% RSLogix 500 project MILLIH2O.RSS, saved by version 12.00.00.00 %
PROJECT "MILLIH2O"    % processor: MicroLogix 1400 %

PROGRAM FILES
  LAD 2   13 rungs
  LAD 3   41 rungs
  LAD 4   59 rungs
  LAD 5   7 rungs
  LAD 6   5 rungs
  LAD 7   8 rungs
  LAD 8   86 rungs

DATA FILES
  O0 OUTPUT  8 elements
  I1 INPUT  8 elements
  S2 STATUS  66 elements
  B3 BINARY  20 elements
  T4 TIMER  27 elements
  C5 COUNTER  11 elements
  R6 CONTROL  1 elements
  N7 INTEGER  50 elements
  F8 FLOAT  133 elements
  N9   17 elements
  F10   3 elements
  B11   5 elements
  F12   23 elements
  N13   50 elements
  N14   4 elements
  C15   10 elements
  C16   10 elements
  B17   4 elements
  F18   60 elements
  F19   10 elements
  N20   100 elements
  B25   1 elements
  B26   1 elements
  F28   10 elements

LADDER 2
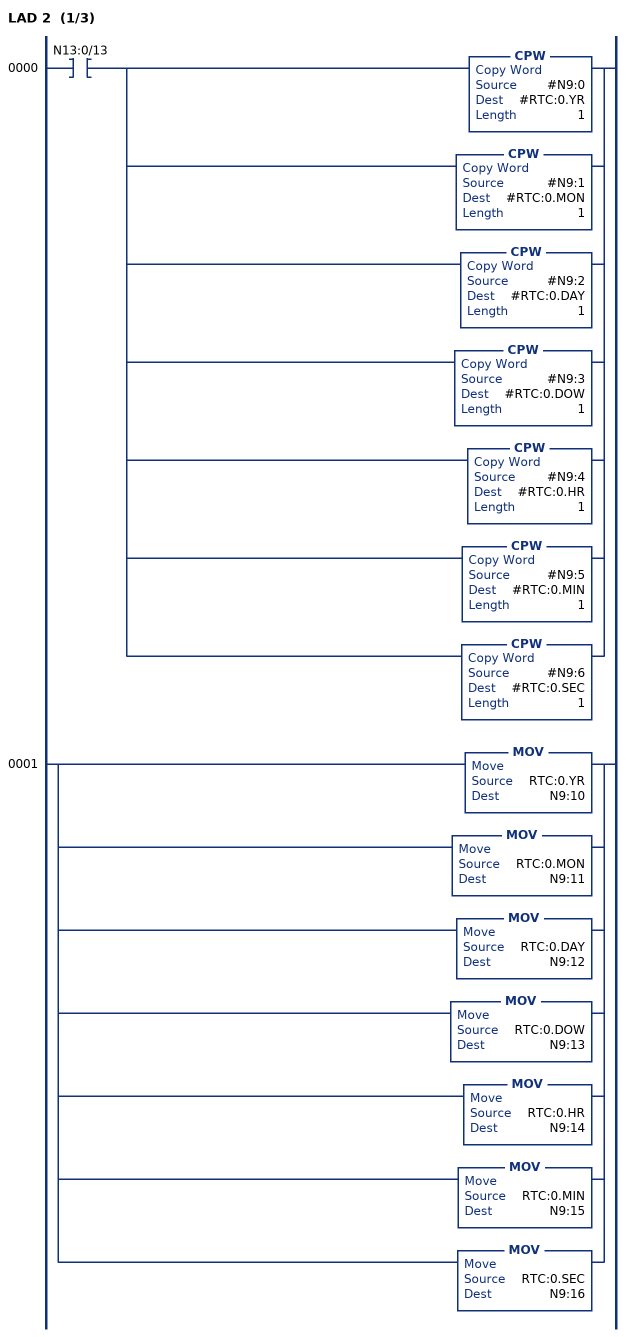
% Rung: 0 %
SOR XIC N13:0/13 BST CPW #N9:0 #RTC:0.YR 1 NXB CPW #N9:1 #RTC:0.MON 1 NXB CPW #N9:2 #RTC:0.DAY 1 NXB CPW #N9:3 #RTC:0.DOW 1 NXB CPW #N9:4 #RTC:0.HR 1 NXB CPW #N9:5 #RTC:0.MIN 1 NXB CPW #N9:6 #RTC:0.SEC 1 BND EOR
% Rung: 1 %
SOR BST MOV RTC:0.YR N9:10 NXB MOV RTC:0.MON N9:11 NXB MOV RTC:0.DAY N9:12 NXB MOV RTC:0.DOW N9:13 NXB MOV RTC:0.HR N9:14 NXB MOV RTC:0.MIN N9:15 NXB MOV RTC:0.SEC N9:16 BND EOR

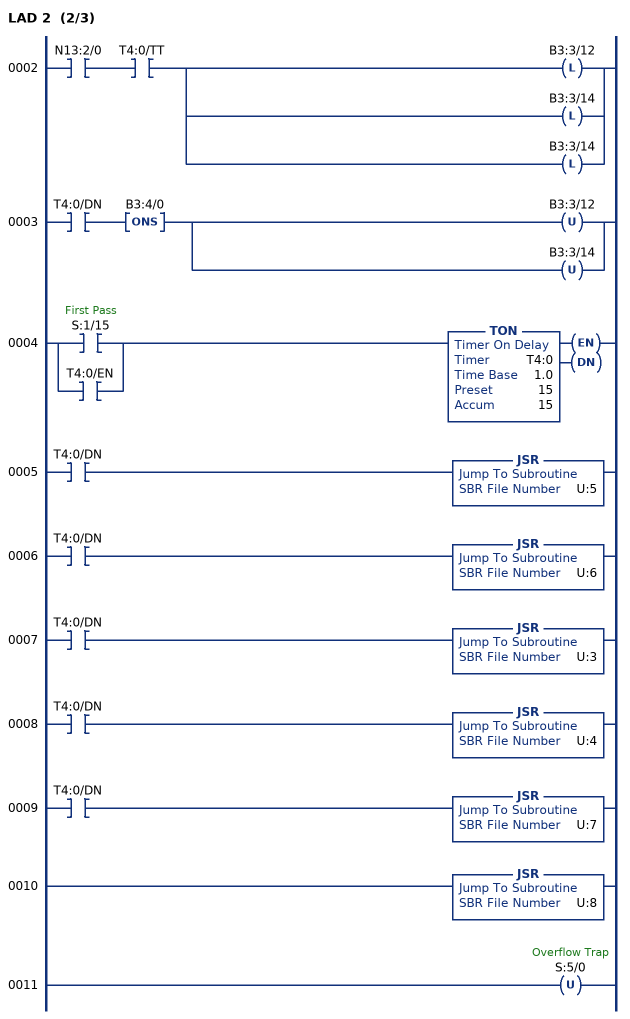
% Rung: 2 %
SOR XIC N13:2/0 XIC T4:0/TT BST OTL B3:3/12 NXB OTL B3:3/14 NXB OTL B3:3/14 BND EOR
% Rung: 3 %
SOR XIC T4:0/DN ONS B3:4/0 BST OTU B3:3/12 NXB OTU B3:3/14 BND EOR
% Rung: 4 %
SOR BST XIC S:1/15 NXB XIC T4:0/EN BND TON T4:0 1.0 15 15 EOR
%   S:1/15  "First Pass" %
% Rung: 5 %
SOR XIC T4:0/DN JSR U:5 EOR
% Rung: 6 %
SOR XIC T4:0/DN JSR U:6 EOR
% Rung: 7 %
SOR XIC T4:0/DN JSR U:3 EOR
% Rung: 8 %
SOR XIC T4:0/DN JSR U:4 EOR
% Rung: 9 %
SOR XIC T4:0/DN JSR U:7 EOR
% Rung: 10 %
SOR JSR U:8 EOR
% Rung: 11 %
SOR OTU S:5/0 EOR
%   S:5/0  "Overflow Trap" %

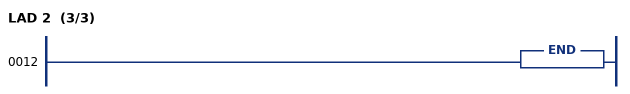
% Rung: 12 %
SOR END EOR

LADDER 3
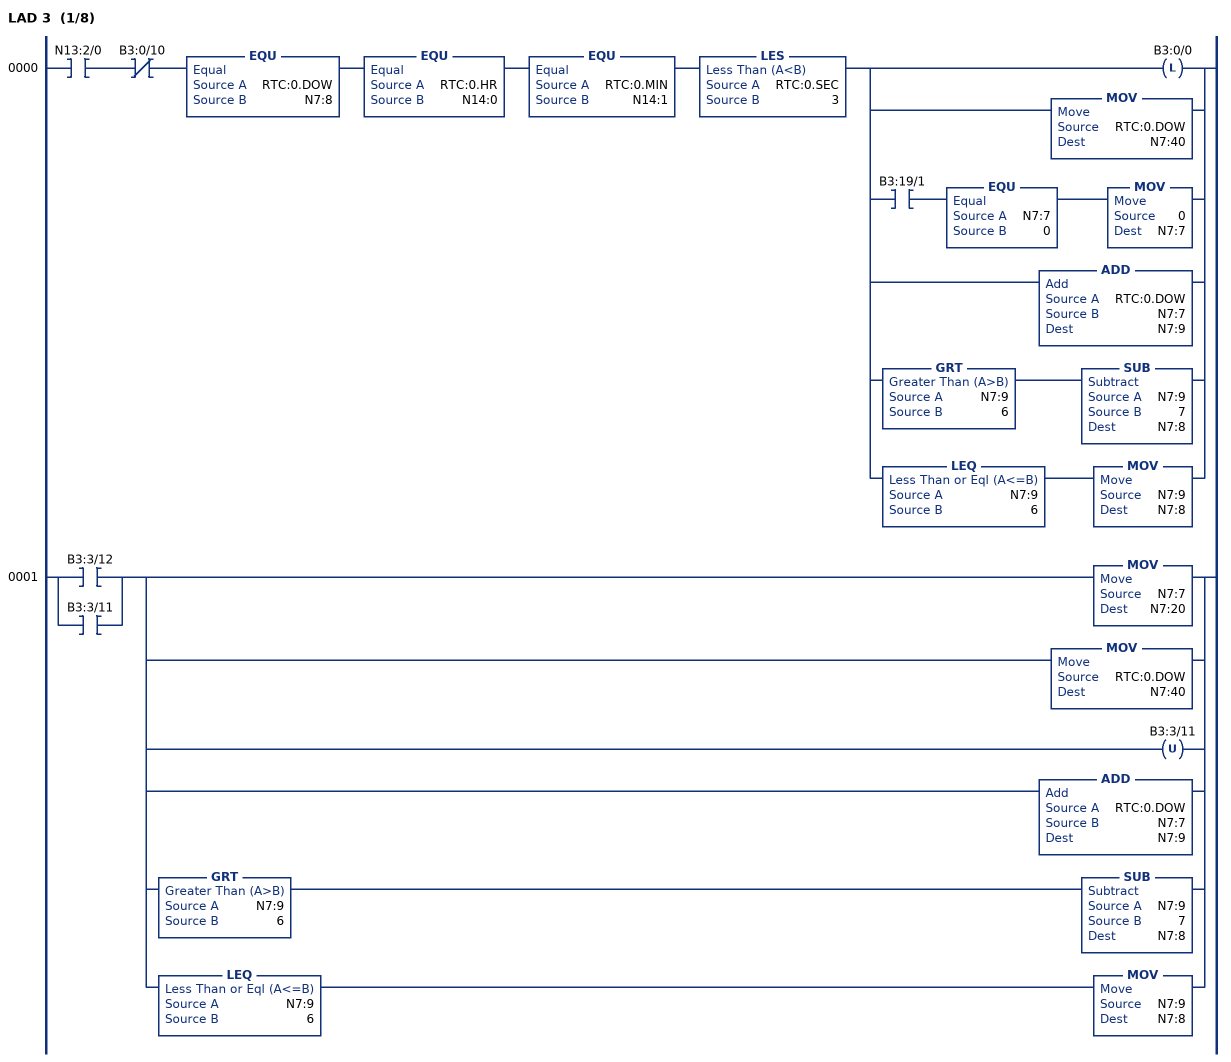
% Rung: 0 %
SOR XIC N13:2/0 XIO B3:0/10 EQU RTC:0.DOW N7:8 EQU RTC:0.HR N14:0 EQU RTC:0.MIN N14:1 LES RTC:0.SEC 3 BST OTL B3:0/0 NXB MOV RTC:0.DOW N7:40 NXB XIC B3:19/1 EQU N7:7 0 MOV 0 N7:7 NXB ADD RTC:0.DOW N7:7 N7:9 NXB GRT N7:9 6 SUB N7:9 7 N7:8 NXB LEQ N7:9 6 MOV N7:9 N7:8 BND EOR
% Rung: 1 %
SOR BST XIC B3:3/12 NXB XIC B3:3/11 BND BST MOV N7:7 N7:20 NXB MOV RTC:0.DOW N7:40 NXB OTU B3:3/11 NXB ADD RTC:0.DOW N7:7 N7:9 NXB GRT N7:9 6 SUB N7:9 7 N7:8 NXB LEQ N7:9 6 MOV N7:9 N7:8 BND EOR

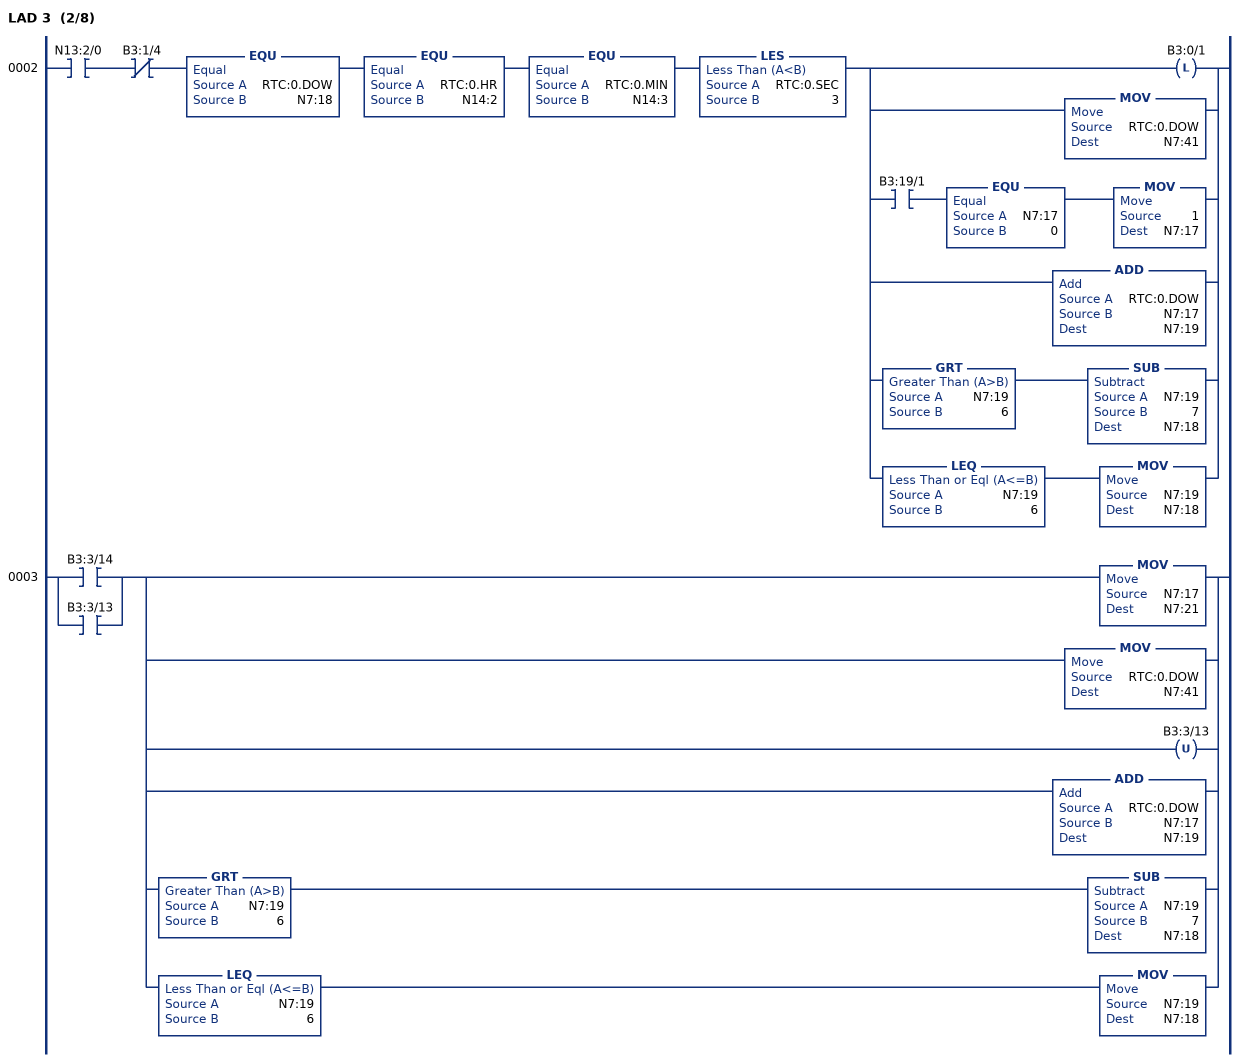
% Rung: 2 %
SOR XIC N13:2/0 XIO B3:1/4 EQU RTC:0.DOW N7:18 EQU RTC:0.HR N14:2 EQU RTC:0.MIN N14:3 LES RTC:0.SEC 3 BST OTL B3:0/1 NXB MOV RTC:0.DOW N7:41 NXB XIC B3:19/1 EQU N7:17 0 MOV 1 N7:17 NXB ADD RTC:0.DOW N7:17 N7:19 NXB GRT N7:19 6 SUB N7:19 7 N7:18 NXB LEQ N7:19 6 MOV N7:19 N7:18 BND EOR
% Rung: 3 %
SOR BST XIC B3:3/14 NXB XIC B3:3/13 BND BST MOV N7:17 N7:21 NXB MOV RTC:0.DOW N7:41 NXB OTU B3:3/13 NXB ADD RTC:0.DOW N7:17 N7:19 NXB GRT N7:19 6 SUB N7:19 7 N7:18 NXB LEQ N7:19 6 MOV N7:19 N7:18 BND EOR

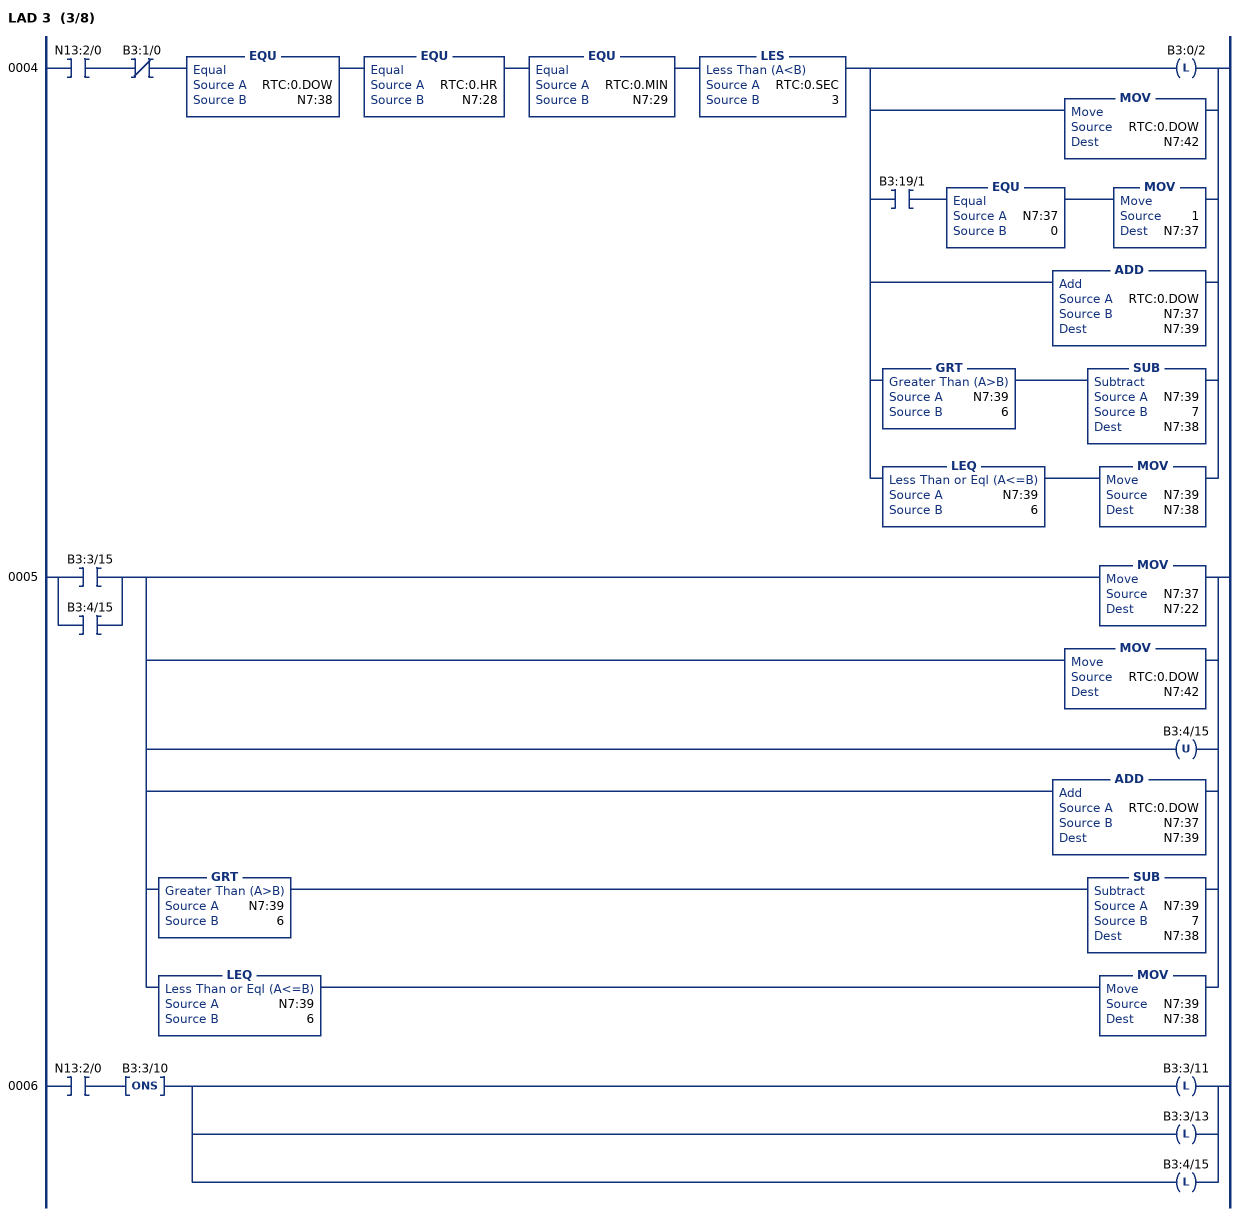
% Rung: 4 %
SOR XIC N13:2/0 XIO B3:1/0 EQU RTC:0.DOW N7:38 EQU RTC:0.HR N7:28 EQU RTC:0.MIN N7:29 LES RTC:0.SEC 3 BST OTL B3:0/2 NXB MOV RTC:0.DOW N7:42 NXB XIC B3:19/1 EQU N7:37 0 MOV 1 N7:37 NXB ADD RTC:0.DOW N7:37 N7:39 NXB GRT N7:39 6 SUB N7:39 7 N7:38 NXB LEQ N7:39 6 MOV N7:39 N7:38 BND EOR
% Rung: 5 %
SOR BST XIC B3:3/15 NXB XIC B3:4/15 BND BST MOV N7:37 N7:22 NXB MOV RTC:0.DOW N7:42 NXB OTU B3:4/15 NXB ADD RTC:0.DOW N7:37 N7:39 NXB GRT N7:39 6 SUB N7:39 7 N7:38 NXB LEQ N7:39 6 MOV N7:39 N7:38 BND EOR
% Rung: 6 %
SOR XIC N13:2/0 ONS B3:3/10 BST OTL B3:3/11 NXB OTL B3:3/13 NXB OTL B3:4/15 BND EOR

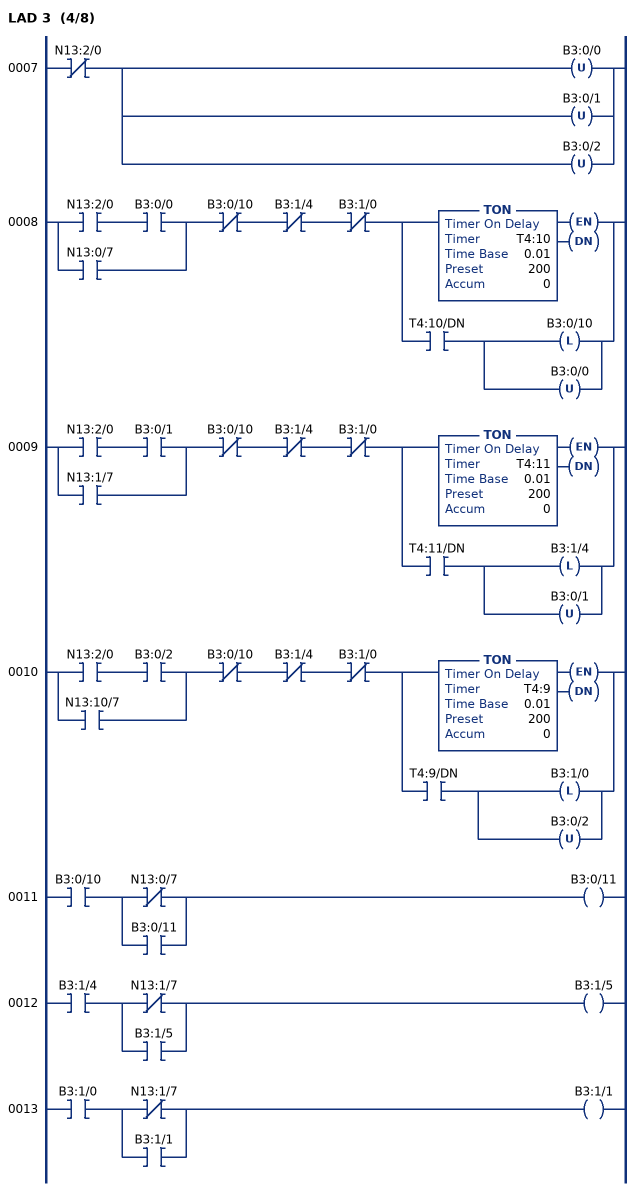
% Rung: 7 %
SOR XIO N13:2/0 BST OTU B3:0/0 NXB OTU B3:0/1 NXB OTU B3:0/2 BND EOR
% Rung: 8 %
SOR BST XIC N13:2/0 XIC B3:0/0 NXB XIC N13:0/7 BND XIO B3:0/10 XIO B3:1/4 XIO B3:1/0 BST TON T4:10 0.01 200 0 NXB XIC T4:10/DN BST OTL B3:0/10 NXB OTU B3:0/0 BND BND EOR
% Rung: 9 %
SOR BST XIC N13:2/0 XIC B3:0/1 NXB XIC N13:1/7 BND XIO B3:0/10 XIO B3:1/4 XIO B3:1/0 BST TON T4:11 0.01 200 0 NXB XIC T4:11/DN BST OTL B3:1/4 NXB OTU B3:0/1 BND BND EOR
% Rung: 10 %
SOR BST XIC N13:2/0 XIC B3:0/2 NXB XIC N13:10/7 BND XIO B3:0/10 XIO B3:1/4 XIO B3:1/0 BST TON T4:9 0.01 200 0 NXB XIC T4:9/DN BST OTL B3:1/0 NXB OTU B3:0/2 BND BND EOR
% Rung: 11 %
SOR XIC B3:0/10 BST XIO N13:0/7 NXB XIC B3:0/11 BND OTE B3:0/11 EOR
% Rung: 12 %
SOR XIC B3:1/4 BST XIO N13:1/7 NXB XIC B3:1/5 BND OTE B3:1/5 EOR
% Rung: 13 %
SOR XIC B3:1/0 BST XIO N13:1/7 NXB XIC B3:1/1 BND OTE B3:1/1 EOR

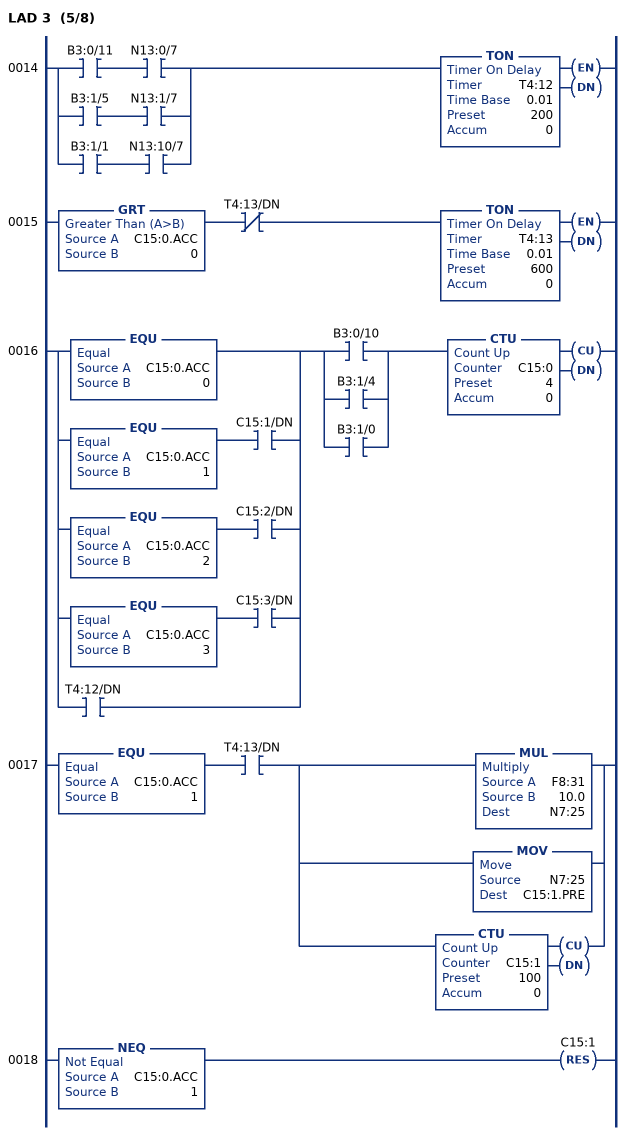
% Rung: 14 %
SOR BST XIC B3:0/11 XIC N13:0/7 NXB XIC B3:1/5 XIC N13:1/7 NXB XIC B3:1/1 XIC N13:10/7 BND TON T4:12 0.01 200 0 EOR
% Rung: 15 %
SOR GRT C15:0.ACC 0 XIO T4:13/DN TON T4:13 0.01 600 0 EOR
% Rung: 16 %
SOR BST EQU C15:0.ACC 0 NXB EQU C15:0.ACC 1 XIC C15:1/DN NXB EQU C15:0.ACC 2 XIC C15:2/DN NXB EQU C15:0.ACC 3 XIC C15:3/DN NXB XIC T4:12/DN BND BST XIC B3:0/10 NXB XIC B3:1/4 NXB XIC B3:1/0 BND CTU C15:0 4 0 EOR
% Rung: 17 %
SOR EQU C15:0.ACC 1 XIC T4:13/DN BST MUL F8:31 10.0 N7:25 NXB MOV N7:25 C15:1.PRE NXB CTU C15:1 100 0 BND EOR
% Rung: 18 %
SOR NEQ C15:0.ACC 1 RES C15:1 EOR

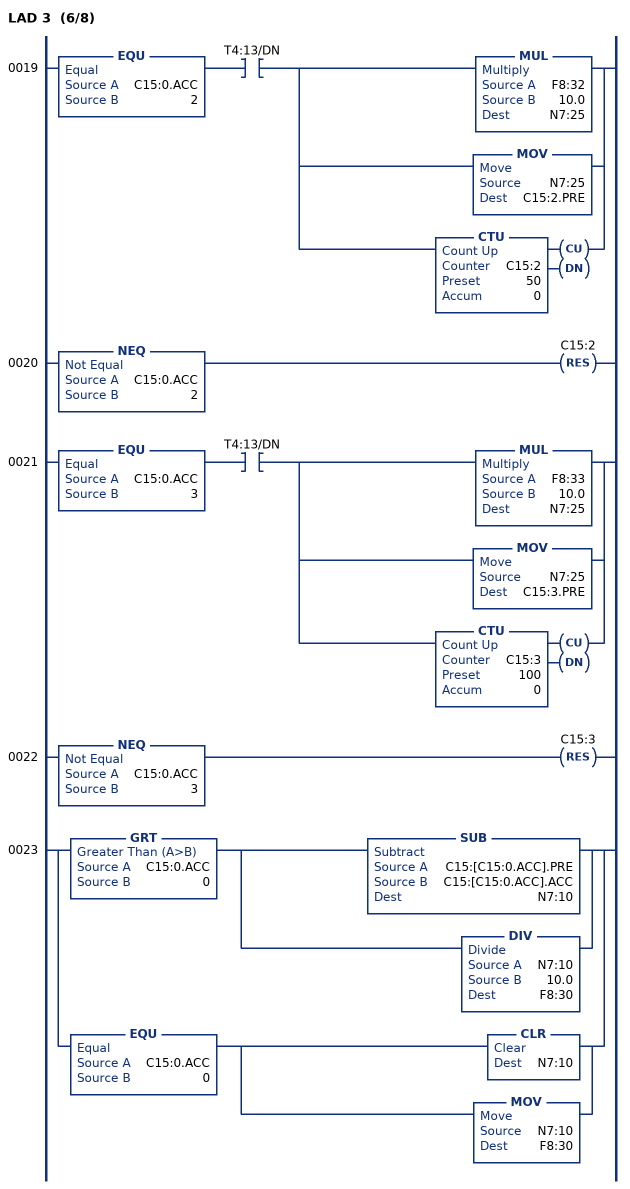
% Rung: 19 %
SOR EQU C15:0.ACC 2 XIC T4:13/DN BST MUL F8:32 10.0 N7:25 NXB MOV N7:25 C15:2.PRE NXB CTU C15:2 50 0 BND EOR
% Rung: 20 %
SOR NEQ C15:0.ACC 2 RES C15:2 EOR
% Rung: 21 %
SOR EQU C15:0.ACC 3 XIC T4:13/DN BST MUL F8:33 10.0 N7:25 NXB MOV N7:25 C15:3.PRE NXB CTU C15:3 100 0 BND EOR
% Rung: 22 %
SOR NEQ C15:0.ACC 3 RES C15:3 EOR
% Rung: 23 %
SOR BST GRT C15:0.ACC 0 BST SUB C15:[C15:0.ACC].PRE C15:[C15:0.ACC].ACC N7:10 NXB DIV N7:10 10.0 F8:30 BND NXB EQU C15:0.ACC 0 BST CLR N7:10 NXB MOV N7:10 F8:30 BND BND EOR

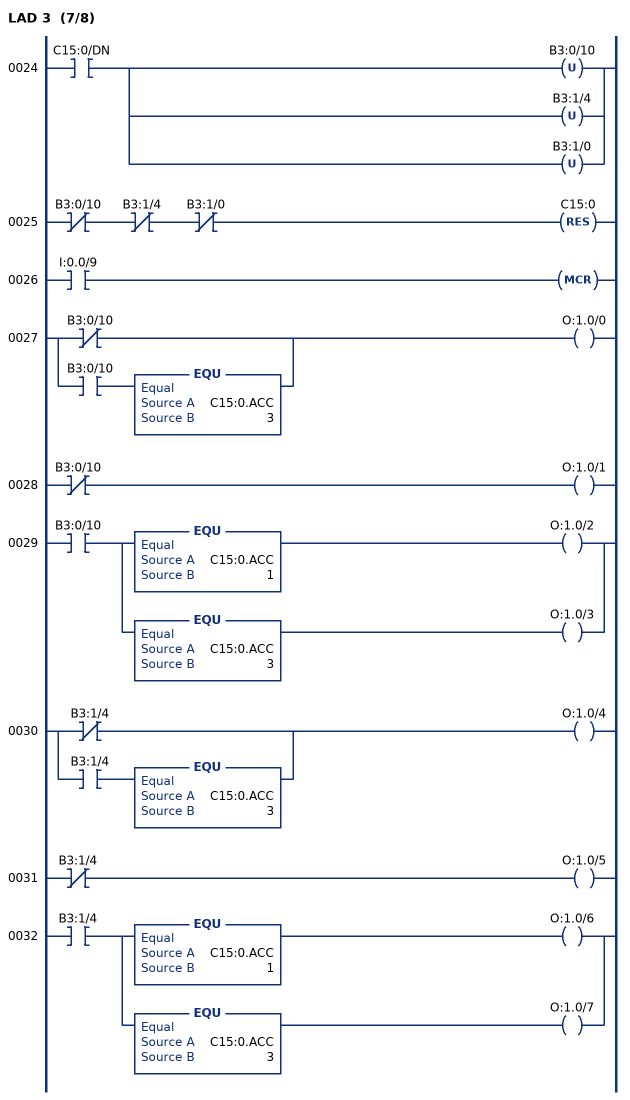
% Rung: 24 %
SOR XIC C15:0/DN BST OTU B3:0/10 NXB OTU B3:1/4 NXB OTU B3:1/0 BND EOR
% Rung: 25 %
SOR XIO B3:0/10 XIO B3:1/4 XIO B3:1/0 RES C15:0 EOR
% Rung: 26 %
SOR XIC I:0.0/9 MCR EOR
% Rung: 27 %
SOR BST XIO B3:0/10 NXB XIC B3:0/10 EQU C15:0.ACC 3 BND OTE O:1.0/0 EOR
% Rung: 28 %
SOR XIO B3:0/10 OTE O:1.0/1 EOR
% Rung: 29 %
SOR XIC B3:0/10 BST EQU C15:0.ACC 1 OTE O:1.0/2 NXB EQU C15:0.ACC 3 OTE O:1.0/3 BND EOR
% Rung: 30 %
SOR BST XIO B3:1/4 NXB XIC B3:1/4 EQU C15:0.ACC 3 BND OTE O:1.0/4 EOR
% Rung: 31 %
SOR XIO B3:1/4 OTE O:1.0/5 EOR
% Rung: 32 %
SOR XIC B3:1/4 BST EQU C15:0.ACC 1 OTE O:1.0/6 NXB EQU C15:0.ACC 3 OTE O:1.0/7 BND EOR

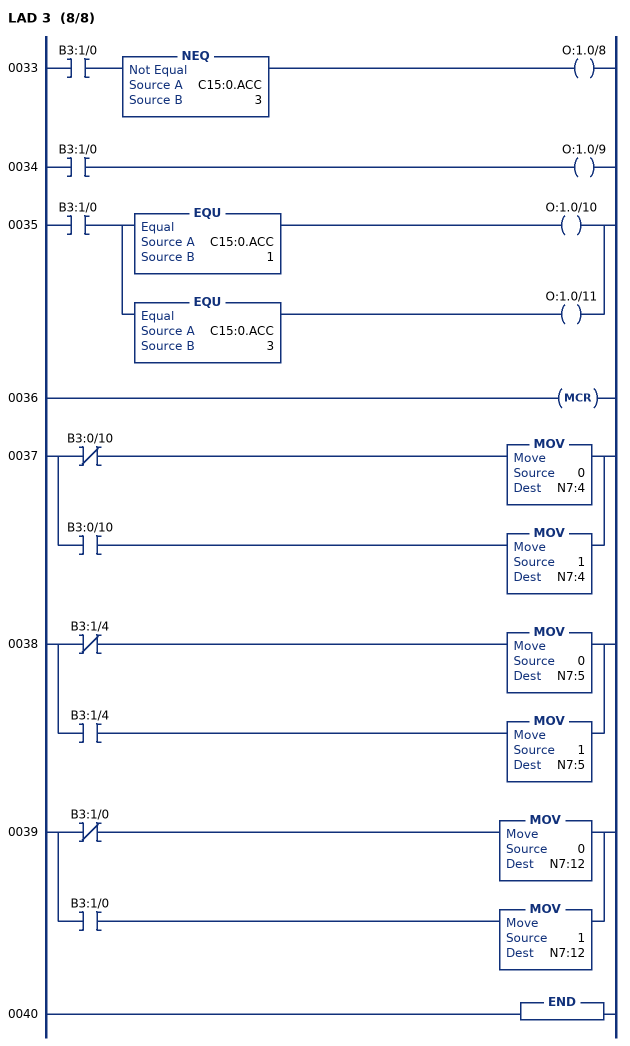
% Rung: 33 %
SOR XIC B3:1/0 NEQ C15:0.ACC 3 OTE O:1.0/8 EOR
% Rung: 34 %
SOR XIC B3:1/0 OTE O:1.0/9 EOR
% Rung: 35 %
SOR XIC B3:1/0 BST EQU C15:0.ACC 1 OTE O:1.0/10 NXB EQU C15:0.ACC 3 OTE O:1.0/11 BND EOR
% Rung: 36 %
SOR MCR EOR
% Rung: 37 %
SOR BST XIO B3:0/10 MOV 0 N7:4 NXB XIC B3:0/10 MOV 1 N7:4 BND EOR
% Rung: 38 %
SOR BST XIO B3:1/4 MOV 0 N7:5 NXB XIC B3:1/4 MOV 1 N7:5 BND EOR
% Rung: 39 %
SOR BST XIO B3:1/0 MOV 0 N7:12 NXB XIC B3:1/0 MOV 1 N7:12 BND EOR
% Rung: 40 %
SOR END EOR

LADDER 4
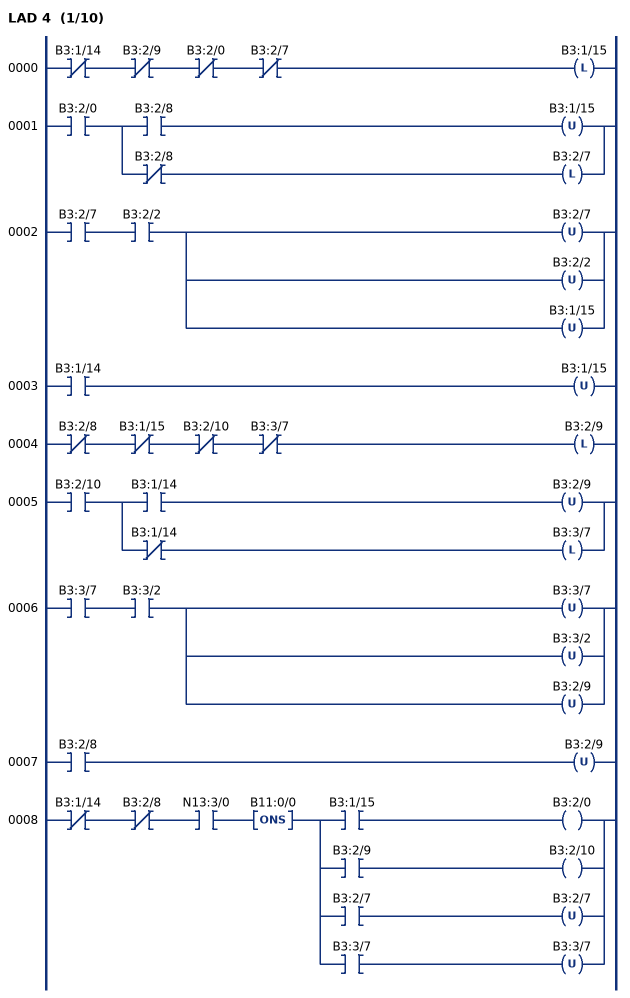
% Rung: 0 %
SOR XIO B3:1/14 XIO B3:2/9 XIO B3:2/0 XIO B3:2/7 OTL B3:1/15 EOR
% Rung: 1 %
SOR XIC B3:2/0 BST XIC B3:2/8 OTU B3:1/15 NXB XIO B3:2/8 OTL B3:2/7 BND EOR
% Rung: 2 %
SOR XIC B3:2/7 XIC B3:2/2 BST OTU B3:2/7 NXB OTU B3:2/2 NXB OTU B3:1/15 BND EOR
% Rung: 3 %
SOR XIC B3:1/14 OTU B3:1/15 EOR
% Rung: 4 %
SOR XIO B3:2/8 XIO B3:1/15 XIO B3:2/10 XIO B3:3/7 OTL B3:2/9 EOR
% Rung: 5 %
SOR XIC B3:2/10 BST XIC B3:1/14 OTU B3:2/9 NXB XIO B3:1/14 OTL B3:3/7 BND EOR
% Rung: 6 %
SOR XIC B3:3/7 XIC B3:3/2 BST OTU B3:3/7 NXB OTU B3:3/2 NXB OTU B3:2/9 BND EOR
% Rung: 7 %
SOR XIC B3:2/8 OTU B3:2/9 EOR
% Rung: 8 %
SOR XIO B3:1/14 XIO B3:2/8 XIC N13:3/0 ONS B11:0/0 BST XIC B3:1/15 OTE B3:2/0 NXB XIC B3:2/9 OTE B3:2/10 NXB XIC B3:2/7 OTU B3:2/7 NXB XIC B3:3/7 OTU B3:3/7 BND EOR

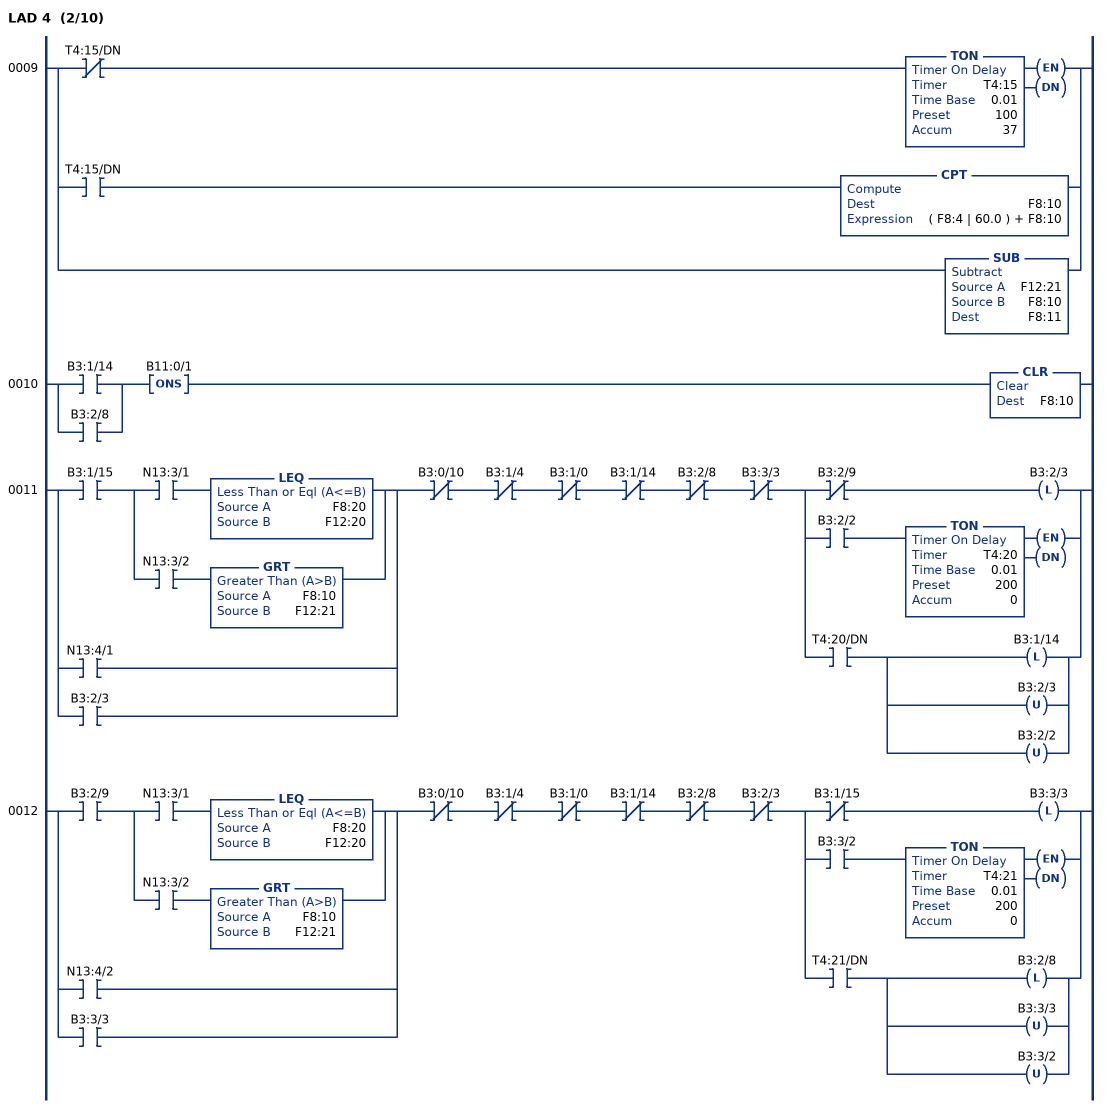
% Rung: 9 %
SOR BST XIO T4:15/DN TON T4:15 0.01 100 37 NXB XIC T4:15/DN CPT F8:10 " ( F8:4 | 60.0 ) + F8:10 " NXB SUB F12:21 F8:10 F8:11 BND EOR
% Rung: 10 %
SOR BST XIC B3:1/14 NXB XIC B3:2/8 BND ONS B11:0/1 CLR F8:10 EOR
% Rung: 11 %
SOR BST XIC B3:1/15 BST XIC N13:3/1 LEQ F8:20 F12:20 NXB XIC N13:3/2 GRT F8:10 F12:21 BND NXB XIC N13:4/1 NXB XIC B3:2/3 BND XIO B3:0/10 XIO B3:1/4 XIO B3:1/0 XIO B3:1/14 XIO B3:2/8 XIO B3:3/3 BST XIO B3:2/9 OTL B3:2/3 NXB XIC B3:2/2 TON T4:20 0.01 200 0 NXB XIC T4:20/DN BST OTL B3:1/14 NXB OTU B3:2/3 NXB OTU B3:2/2 BND BND EOR
% Rung: 12 %
SOR BST XIC B3:2/9 BST XIC N13:3/1 LEQ F8:20 F12:20 NXB XIC N13:3/2 GRT F8:10 F12:21 BND NXB XIC N13:4/2 NXB XIC B3:3/3 BND XIO B3:0/10 XIO B3:1/4 XIO B3:1/0 XIO B3:1/14 XIO B3:2/8 XIO B3:2/3 BST XIO B3:1/15 OTL B3:3/3 NXB XIC B3:3/2 TON T4:21 0.01 200 0 NXB XIC T4:21/DN BST OTL B3:2/8 NXB OTU B3:3/3 NXB OTU B3:3/2 BND BND EOR

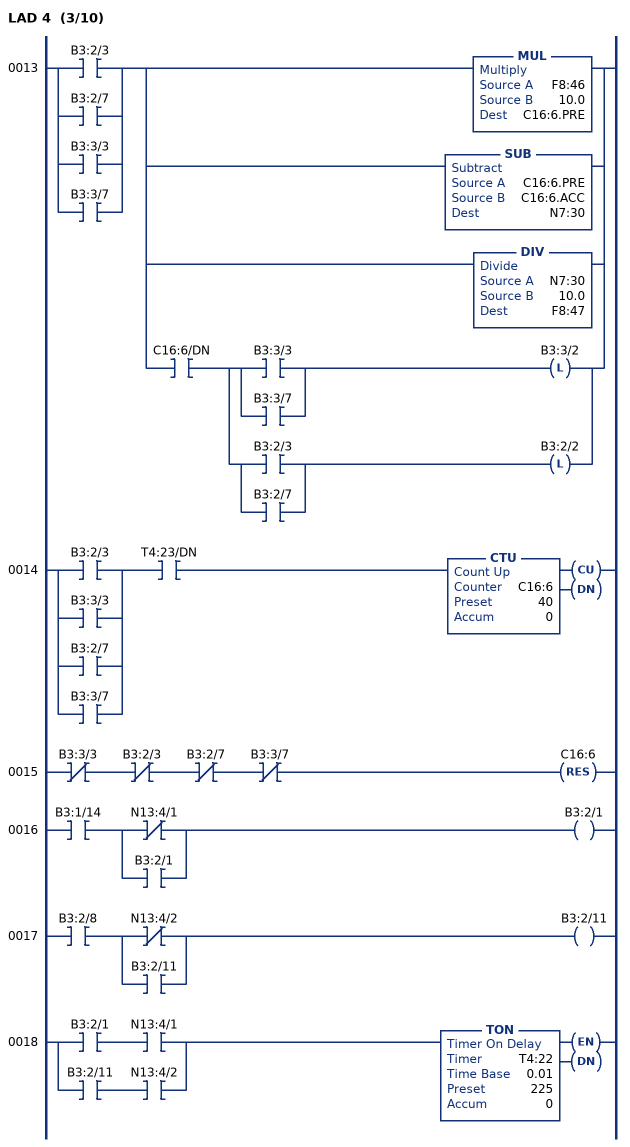
% Rung: 13 %
SOR BST XIC B3:2/3 NXB XIC B3:2/7 NXB XIC B3:3/3 NXB XIC B3:3/7 BND BST MUL F8:46 10.0 C16:6.PRE NXB SUB C16:6.PRE C16:6.ACC N7:30 NXB DIV N7:30 10.0 F8:47 NXB XIC C16:6/DN BST BST XIC B3:3/3 NXB XIC B3:3/7 BND OTL B3:3/2 NXB BST XIC B3:2/3 NXB XIC B3:2/7 BND OTL B3:2/2 BND BND EOR
% Rung: 14 %
SOR BST XIC B3:2/3 NXB XIC B3:3/3 NXB XIC B3:2/7 NXB XIC B3:3/7 BND XIC T4:23/DN CTU C16:6 40 0 EOR
% Rung: 15 %
SOR XIO B3:3/3 XIO B3:2/3 XIO B3:2/7 XIO B3:3/7 RES C16:6 EOR
% Rung: 16 %
SOR XIC B3:1/14 BST XIO N13:4/1 NXB XIC B3:2/1 BND OTE B3:2/1 EOR
% Rung: 17 %
SOR XIC B3:2/8 BST XIO N13:4/2 NXB XIC B3:2/11 BND OTE B3:2/11 EOR
% Rung: 18 %
SOR BST XIC B3:2/1 XIC N13:4/1 NXB XIC B3:2/11 XIC N13:4/2 BND TON T4:22 0.01 225 0 EOR

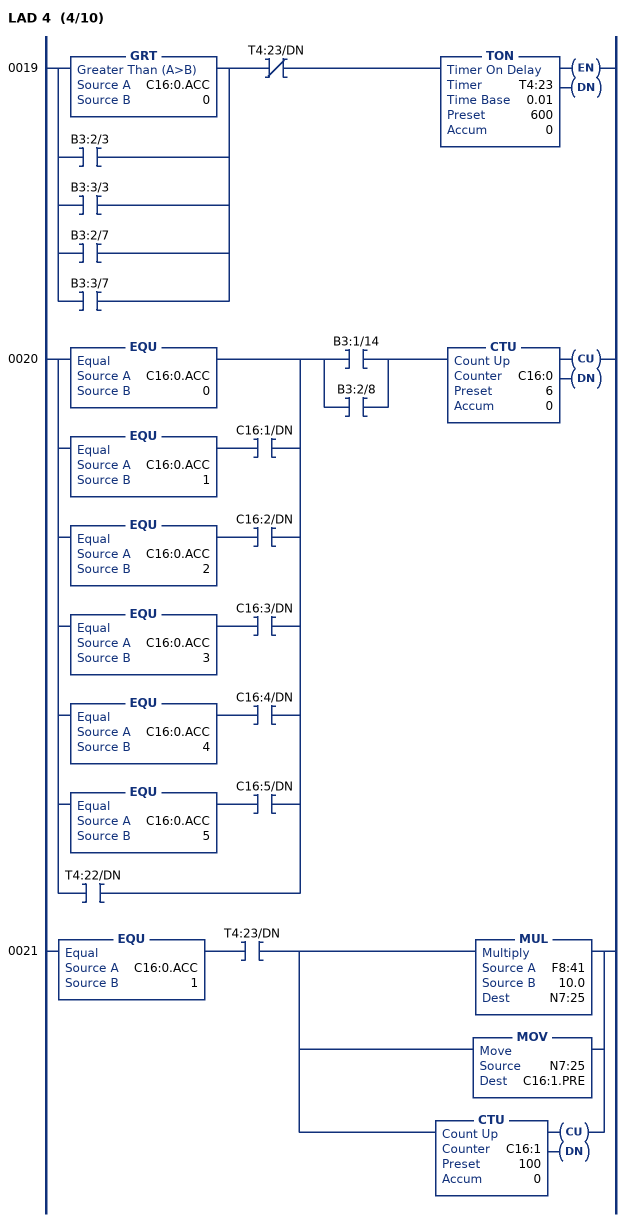
% Rung: 19 %
SOR BST GRT C16:0.ACC 0 NXB XIC B3:2/3 NXB XIC B3:3/3 NXB XIC B3:2/7 NXB XIC B3:3/7 BND XIO T4:23/DN TON T4:23 0.01 600 0 EOR
% Rung: 20 %
SOR BST EQU C16:0.ACC 0 NXB EQU C16:0.ACC 1 XIC C16:1/DN NXB EQU C16:0.ACC 2 XIC C16:2/DN NXB EQU C16:0.ACC 3 XIC C16:3/DN NXB EQU C16:0.ACC 4 XIC C16:4/DN NXB EQU C16:0.ACC 5 XIC C16:5/DN NXB XIC T4:22/DN BND BST XIC B3:1/14 NXB XIC B3:2/8 BND CTU C16:0 6 0 EOR
% Rung: 21 %
SOR EQU C16:0.ACC 1 XIC T4:23/DN BST MUL F8:41 10.0 N7:25 NXB MOV N7:25 C16:1.PRE NXB CTU C16:1 100 0 BND EOR

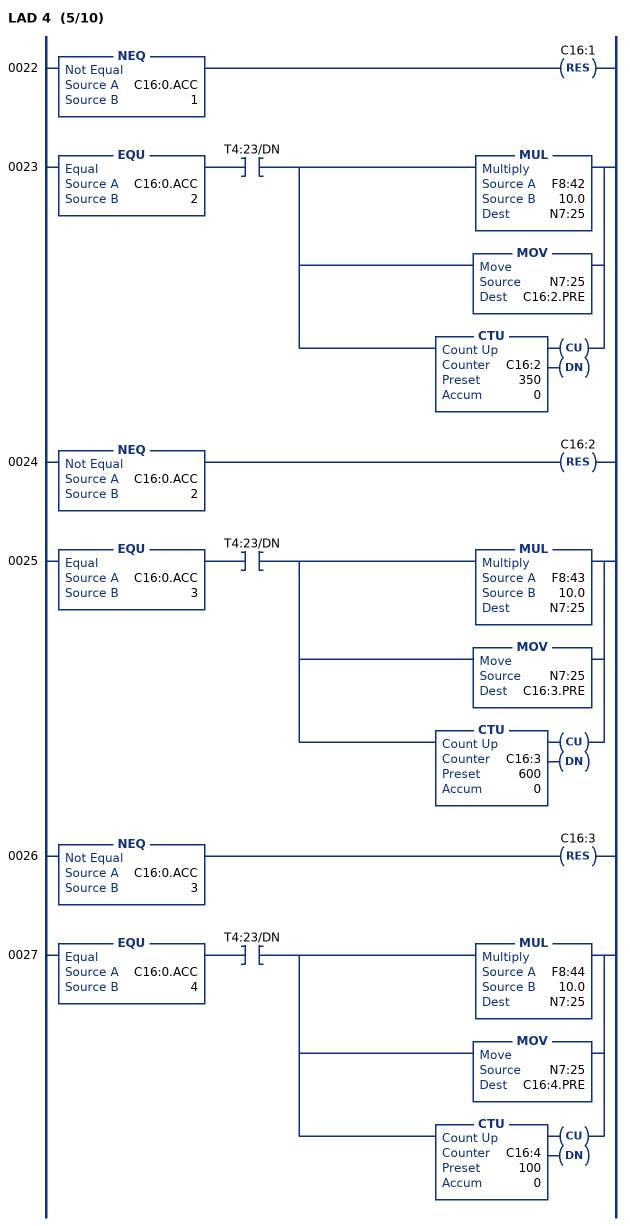
% Rung: 22 %
SOR NEQ C16:0.ACC 1 RES C16:1 EOR
% Rung: 23 %
SOR EQU C16:0.ACC 2 XIC T4:23/DN BST MUL F8:42 10.0 N7:25 NXB MOV N7:25 C16:2.PRE NXB CTU C16:2 350 0 BND EOR
% Rung: 24 %
SOR NEQ C16:0.ACC 2 RES C16:2 EOR
% Rung: 25 %
SOR EQU C16:0.ACC 3 XIC T4:23/DN BST MUL F8:43 10.0 N7:25 NXB MOV N7:25 C16:3.PRE NXB CTU C16:3 600 0 BND EOR
% Rung: 26 %
SOR NEQ C16:0.ACC 3 RES C16:3 EOR
% Rung: 27 %
SOR EQU C16:0.ACC 4 XIC T4:23/DN BST MUL F8:44 10.0 N7:25 NXB MOV N7:25 C16:4.PRE NXB CTU C16:4 100 0 BND EOR

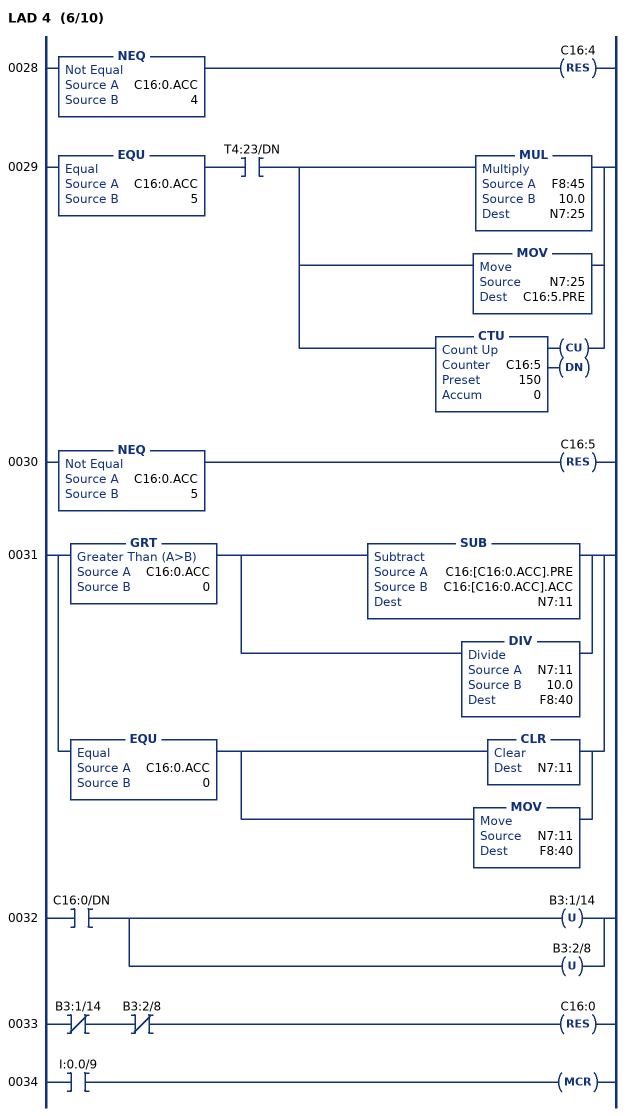
% Rung: 28 %
SOR NEQ C16:0.ACC 4 RES C16:4 EOR
% Rung: 29 %
SOR EQU C16:0.ACC 5 XIC T4:23/DN BST MUL F8:45 10.0 N7:25 NXB MOV N7:25 C16:5.PRE NXB CTU C16:5 150 0 BND EOR
% Rung: 30 %
SOR NEQ C16:0.ACC 5 RES C16:5 EOR
% Rung: 31 %
SOR BST GRT C16:0.ACC 0 BST SUB C16:[C16:0.ACC].PRE C16:[C16:0.ACC].ACC N7:11 NXB DIV N7:11 10.0 F8:40 BND NXB EQU C16:0.ACC 0 BST CLR N7:11 NXB MOV N7:11 F8:40 BND BND EOR
% Rung: 32 %
SOR XIC C16:0/DN BST OTU B3:1/14 NXB OTU B3:2/8 BND EOR
% Rung: 33 %
SOR XIO B3:1/14 XIO B3:2/8 RES C16:0 EOR
% Rung: 34 %
SOR XIC I:0.0/9 MCR EOR

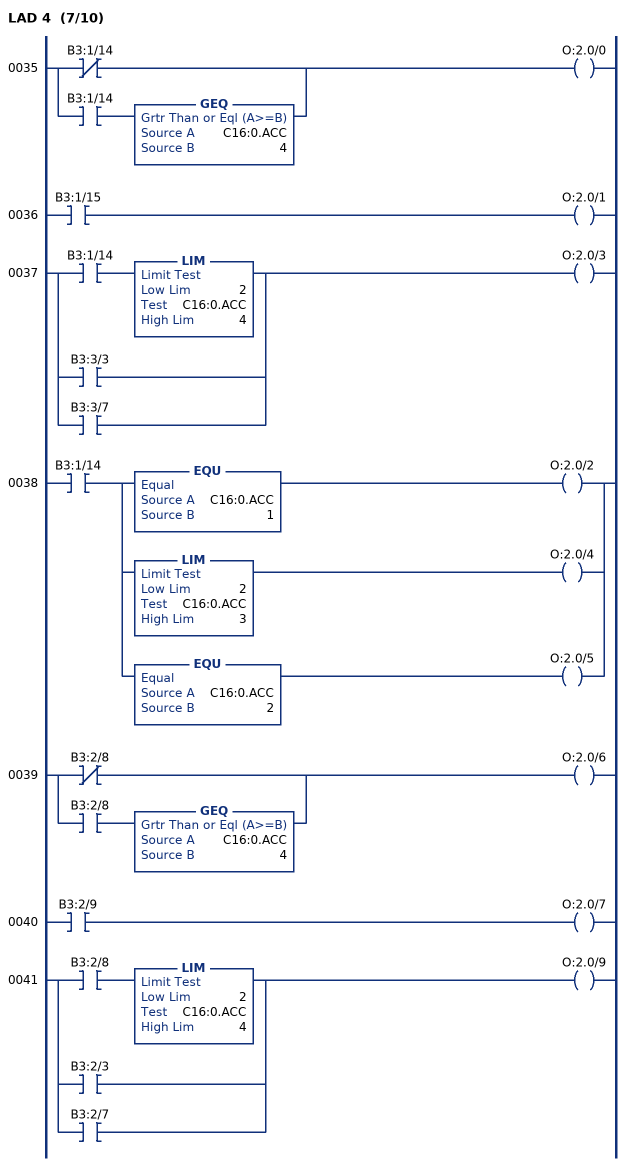
% Rung: 35 %
SOR BST XIO B3:1/14 NXB XIC B3:1/14 GEQ C16:0.ACC 4 BND OTE O:2.0/0 EOR
% Rung: 36 %
SOR XIC B3:1/15 OTE O:2.0/1 EOR
% Rung: 37 %
SOR BST XIC B3:1/14 LIM 2 C16:0.ACC 4 NXB XIC B3:3/3 NXB XIC B3:3/7 BND OTE O:2.0/3 EOR
% Rung: 38 %
SOR XIC B3:1/14 BST EQU C16:0.ACC 1 OTE O:2.0/2 NXB LIM 2 C16:0.ACC 3 OTE O:2.0/4 NXB EQU C16:0.ACC 2 OTE O:2.0/5 BND EOR
% Rung: 39 %
SOR BST XIO B3:2/8 NXB XIC B3:2/8 GEQ C16:0.ACC 4 BND OTE O:2.0/6 EOR
% Rung: 40 %
SOR XIC B3:2/9 OTE O:2.0/7 EOR
% Rung: 41 %
SOR BST XIC B3:2/8 LIM 2 C16:0.ACC 4 NXB XIC B3:2/3 NXB XIC B3:2/7 BND OTE O:2.0/9 EOR

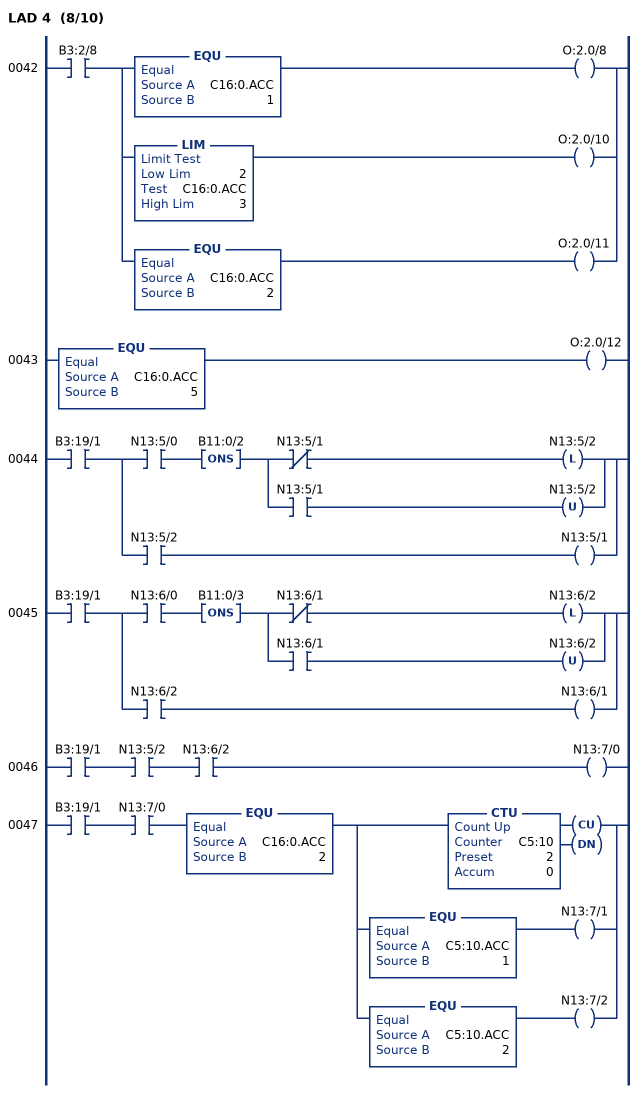
% Rung: 42 %
SOR XIC B3:2/8 BST EQU C16:0.ACC 1 OTE O:2.0/8 NXB LIM 2 C16:0.ACC 3 OTE O:2.0/10 NXB EQU C16:0.ACC 2 OTE O:2.0/11 BND EOR
% Rung: 43 %
SOR EQU C16:0.ACC 5 OTE O:2.0/12 EOR
% Rung: 44 %
SOR XIC B3:19/1 BST XIC N13:5/0 ONS B11:0/2 BST XIO N13:5/1 OTL N13:5/2 NXB XIC N13:5/1 OTU N13:5/2 BND NXB XIC N13:5/2 OTE N13:5/1 BND EOR
% Rung: 45 %
SOR XIC B3:19/1 BST XIC N13:6/0 ONS B11:0/3 BST XIO N13:6/1 OTL N13:6/2 NXB XIC N13:6/1 OTU N13:6/2 BND NXB XIC N13:6/2 OTE N13:6/1 BND EOR
% Rung: 46 %
SOR XIC B3:19/1 XIC N13:5/2 XIC N13:6/2 OTE N13:7/0 EOR
% Rung: 47 %
SOR XIC B3:19/1 XIC N13:7/0 EQU C16:0.ACC 2 BST CTU C5:10 2 0 NXB EQU C5:10.ACC 1 OTE N13:7/1 NXB EQU C5:10.ACC 2 OTE N13:7/2 BND EOR

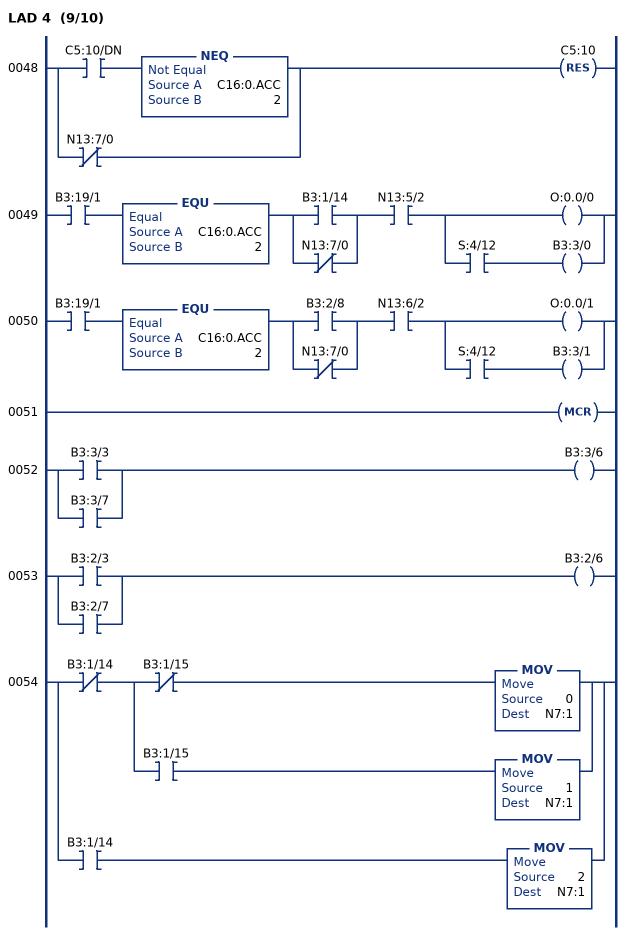
% Rung: 48 %
SOR BST XIC C5:10/DN NEQ C16:0.ACC 2 NXB XIO N13:7/0 BND RES C5:10 EOR
% Rung: 49 %
SOR XIC B3:19/1 EQU C16:0.ACC 2 BST XIC B3:1/14 NXB XIO N13:7/0 BND XIC N13:5/2 BST OTE O:0.0/0 NXB XIC S:4/12 OTE B3:3/0 BND EOR
% Rung: 50 %
SOR XIC B3:19/1 EQU C16:0.ACC 2 BST XIC B3:2/8 NXB XIO N13:7/0 BND XIC N13:6/2 BST OTE O:0.0/1 NXB XIC S:4/12 OTE B3:3/1 BND EOR
% Rung: 51 %
SOR MCR EOR
% Rung: 52 %
SOR BST XIC B3:3/3 NXB XIC B3:3/7 BND OTE B3:3/6 EOR
% Rung: 53 %
SOR BST XIC B3:2/3 NXB XIC B3:2/7 BND OTE B3:2/6 EOR
% Rung: 54 %
SOR BST XIO B3:1/14 BST XIO B3:1/15 MOV 0 N7:1 NXB XIC B3:1/15 MOV 1 N7:1 BND NXB XIC B3:1/14 MOV 2 N7:1 BND EOR

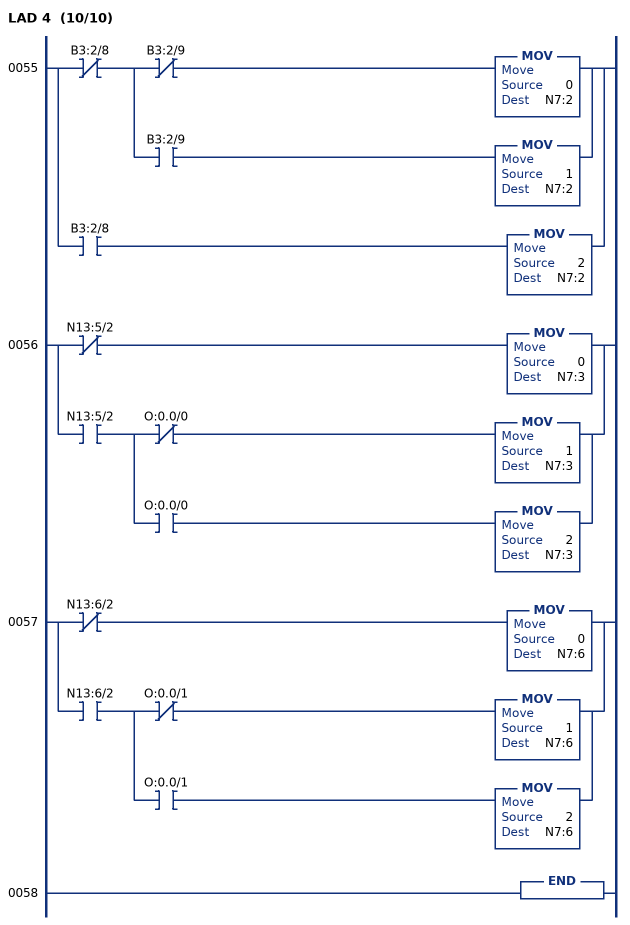
% Rung: 55 %
SOR BST XIO B3:2/8 BST XIO B3:2/9 MOV 0 N7:2 NXB XIC B3:2/9 MOV 1 N7:2 BND NXB XIC B3:2/8 MOV 2 N7:2 BND EOR
% Rung: 56 %
SOR BST XIO N13:5/2 MOV 0 N7:3 NXB XIC N13:5/2 BST XIO O:0.0/0 MOV 1 N7:3 NXB XIC O:0.0/0 MOV 2 N7:3 BND BND EOR
% Rung: 57 %
SOR BST XIO N13:6/2 MOV 0 N7:6 NXB XIC N13:6/2 BST XIO O:0.0/1 MOV 1 N7:6 NXB XIC O:0.0/1 MOV 2 N7:6 BND BND EOR
% Rung: 58 %
SOR END EOR

LADDER 5
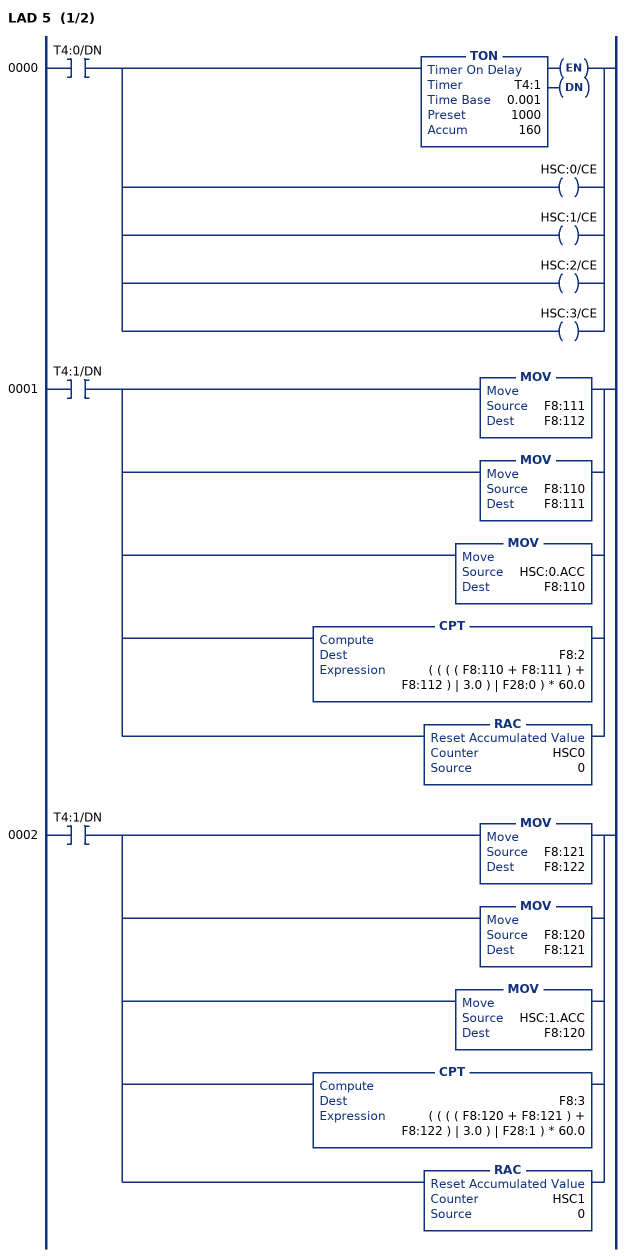
% Rung: 0 %
SOR XIC T4:0/DN BST TON T4:1 0.001 1000 160 NXB OTE HSC:0/CE NXB OTE HSC:1/CE NXB OTE HSC:2/CE NXB OTE HSC:3/CE BND EOR
% Rung: 1 %
SOR XIC T4:1/DN BST MOV F8:111 F8:112 NXB MOV F8:110 F8:111 NXB MOV HSC:0.ACC F8:110 NXB CPT F8:2 " ( ( ( ( F8:110 + F8:111 ) + F8:112 ) | 3.0 ) | F28:0 ) * 60.0 " NXB RAC HSC0 0 BND EOR
% Rung: 2 %
SOR XIC T4:1/DN BST MOV F8:121 F8:122 NXB MOV F8:120 F8:121 NXB MOV HSC:1.ACC F8:120 NXB CPT F8:3 " ( ( ( ( F8:120 + F8:121 ) + F8:122 ) | 3.0 ) | F28:1 ) * 60.0 " NXB RAC HSC1 0 BND EOR

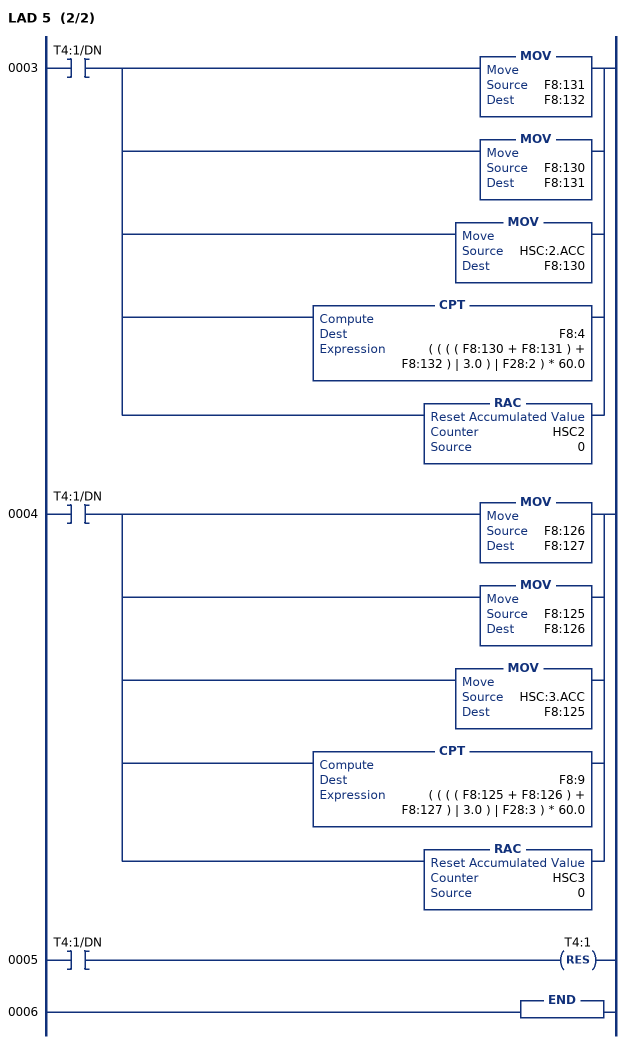
% Rung: 3 %
SOR XIC T4:1/DN BST MOV F8:131 F8:132 NXB MOV F8:130 F8:131 NXB MOV HSC:2.ACC F8:130 NXB CPT F8:4 " ( ( ( ( F8:130 + F8:131 ) + F8:132 ) | 3.0 ) | F28:2 ) * 60.0 " NXB RAC HSC2 0 BND EOR
% Rung: 4 %
SOR XIC T4:1/DN BST MOV F8:126 F8:127 NXB MOV F8:125 F8:126 NXB MOV HSC:3.ACC F8:125 NXB CPT F8:9 " ( ( ( ( F8:125 + F8:126 ) + F8:127 ) | 3.0 ) | F28:3 ) * 60.0 " NXB RAC HSC3 0 BND EOR
% Rung: 5 %
SOR XIC T4:1/DN RES T4:1 EOR
% Rung: 6 %
SOR END EOR

LADDER 6
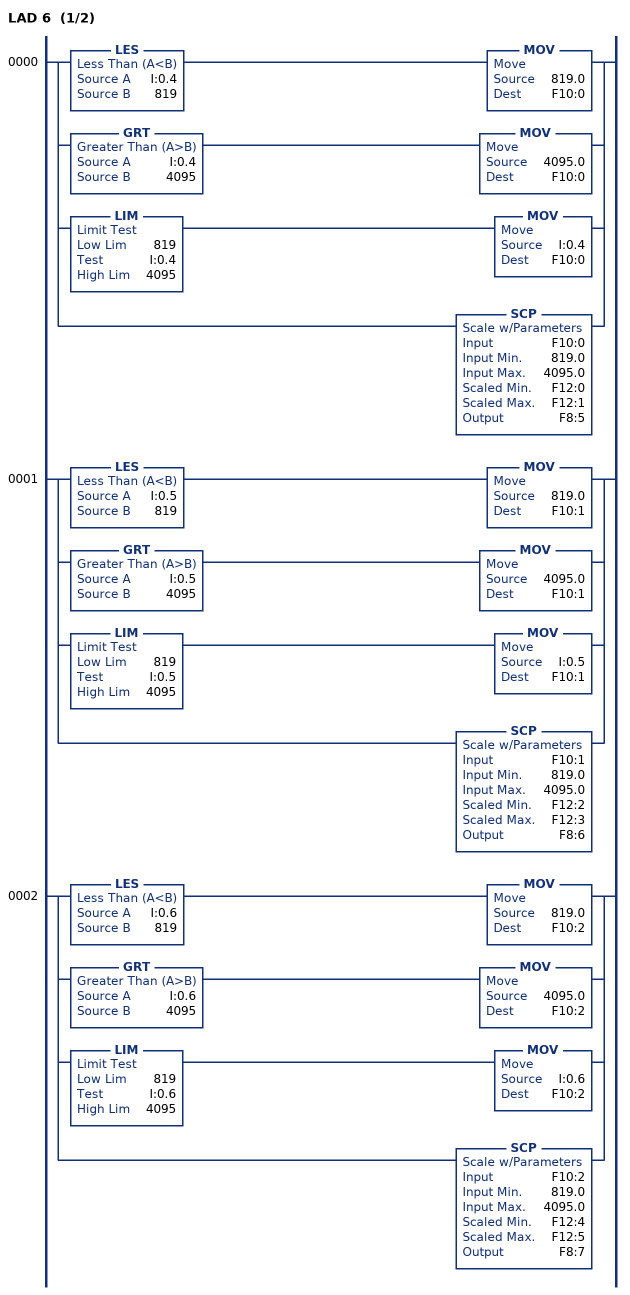
% Rung: 0 %
SOR BST LES I:0.4 819 MOV 819.0 F10:0 NXB GRT I:0.4 4095 MOV 4095.0 F10:0 NXB LIM 819 I:0.4 4095 MOV I:0.4 F10:0 NXB SCP F10:0 819.0 4095.0 F12:0 F12:1 F8:5 BND EOR
% Rung: 1 %
SOR BST LES I:0.5 819 MOV 819.0 F10:1 NXB GRT I:0.5 4095 MOV 4095.0 F10:1 NXB LIM 819 I:0.5 4095 MOV I:0.5 F10:1 NXB SCP F10:1 819.0 4095.0 F12:2 F12:3 F8:6 BND EOR
% Rung: 2 %
SOR BST LES I:0.6 819 MOV 819.0 F10:2 NXB GRT I:0.6 4095 MOV 4095.0 F10:2 NXB LIM 819 I:0.6 4095 MOV I:0.6 F10:2 NXB SCP F10:2 819.0 4095.0 F12:4 F12:5 F8:7 BND EOR

